{attribute 'pack_mode' := '1'}
TYPE ST_BatConfig_Rx :
STRUCT
	DeviceId : UDINT;
	SocMin : REAL;
	SocMax : REAL;
END_STRUCT
END_TYPE

(* stored: Version 1.1.0.1, ProductVersion 3.1.4024.12
   DUT ST_BatConfig_Rx: Id {c5f1ed29-57a2-4544-8b18-b57968d3678a} *)
